(* IEC 61131-3 sources: plcassist-cli/packages/volt-lsp-iec/test-corpus/awa-palletizer/Device/Plc Logic/Application/Library Manager/SysTimeCore, 3 files *)

(* ---- SYSTIMEGETMS.fun ---- *)
FUNCTION SYSTIMEGETMS : UDINT
END_FUNCTION

(* ---- SYSTIMEGETNS.fun ---- *)
FUNCTION SYSTIMEGETNS : RTS_IEC_RESULT
VAR_IN_OUT
	PUSTIME : SYSTIME;
END_VAR
END_FUNCTION

(* ---- SYSTIMEGETUS.fun ---- *)
FUNCTION SYSTIMEGETUS : RTS_IEC_RESULT
VAR_IN_OUT
	PUSTIME : SYSTIME;
END_VAR
END_FUNCTION
